Fanuc KAREL source: kt00994.KL

PROGRAM KT00994
%STACKSIZE=65535
%PRIORITY=65535
%NOLOCKGROUP
VAR
P1 : JOINTPOS9
P2 : JOINTPOS9
X : REAL
Y : REAL
Z : REAL
W : REAL
P : REAL
R : REAL
-- UNRESOLVED DECLARATIONS (source type spelling not recovered)
-- CFG : TYPE_0x001C (type_u16=0x001C)
BEGIN
-- UNRESOLVED_PC line 14 opcodes [27 27 49 7E AD 22 22 22 22 22 22 22 76] marker_code=0
END KT00994
